// Mitsubishi GX Works2 project: 수위제어   PLC: Q02/Q02H

PROGRAM MAIN
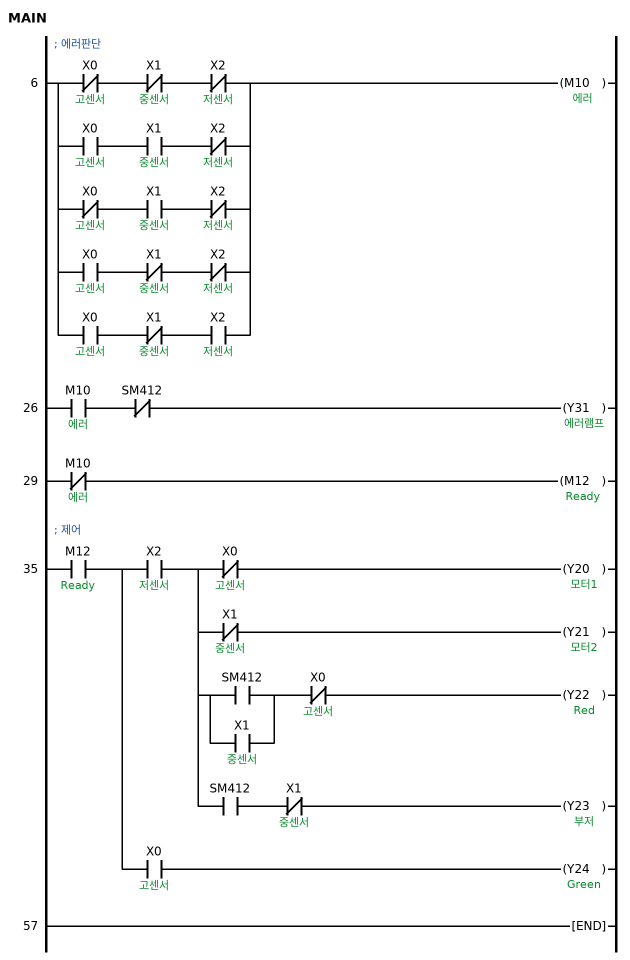
; 에러판단
6     LDI     X0  ; 고센서
      ANI     X1  ; 중센서
      ANI     X2  ; 저센서
      LD      X0  ; 고센서
      AND     X1  ; 중센서
      ANI     X2  ; 저센서
      ORB
      LDI     X0  ; 고센서
      AND     X1  ; 중센서
      ANI     X2  ; 저센서
      ORB
      LD      X0  ; 고센서
      ANI     X1  ; 중센서
      ANI     X2  ; 저센서
      ORB
      LD      X0  ; 고센서
      ANI     X1  ; 중센서
      AND     X2  ; 저센서
      ORB
      OUT     M10  ; 에러
26    LD      M10  ; 에러
      ANI     SM412
      OUT     Y31  ; 에러램프
29    LDI     M10  ; 에러
      OUT     M12  ; Ready
; 제어
35    LD      M12  ; Ready
      MPS
      AND     X2  ; 저센서
      MPS
      ANI     X0  ; 고센서
      OUT     Y20  ; 모터1
      MRD
      ANI     X1  ; 중센서
      OUT     Y21  ; 모터2
      MRD
      LD      SM412
      OR      X1  ; 중센서
      ANB
      ANI     X0  ; 고센서
      OUT     Y22  ; Red
      MPP
      AND     SM412
      ANI     X1  ; 중센서
      OUT     Y23  ; 부저
      MPP
      AND     X0  ; 고센서
      OUT     Y24  ; Green
57    END
END_PROGRAM

// device comments not shown above
X3  ; 테스트
